(* IEC 61131-3 sources: SRCI_CLIENT_PLC/RobotLibrary/Library/POUs/Calculation/MC_CalculateTool/Structures, 4 files *)

(* ---- CalculateToolOutCmd.st ---- *)
{attribute 'pack_mode' := '1'}
// -------------------------------------------------------------------------
//  SRCI Robot Library
// -------------------------------------------------------------------------
//
//  Object:      CalculateToolOutCmd
//  Author:      Thorsten Brach
//  Date:        2024-06-09
//
//  Description:
//
//
//  Copyright:
//    (C) 2024 Thorsten Brach. All rights reserved
//             Licensed under the MIT License.
//
//  Disclaimer:
//    This project is provided without any guarantee and can be used for
//    private and commercial purposes. Any use is at the user’s
//    own risk and responsibility.
//
// -------------------------------------------------------------------------
TYPE CalculateToolOutCmd :
STRUCT
  /// Tool data
  ToolData           : ToolData;
  /// Maximum error of deviation of the TCP position
  /// from the fix point in world coordinate system
  /// If not supported: • -1
  TCPMaxError       : REAL;
  /// Average error of TCP position from the fix point  in world coordinate system
  /// If not supported: • -1
  TCPMeanError      : REAL;
END_STRUCT
END_TYPE

(* ---- CalculateToolParCmd.st ---- *)
{attribute 'pack_mode' := '1'}
// -------------------------------------------------------------------------
//  SRCI Robot Library
// -------------------------------------------------------------------------
//
//  Object:      CalculateToolParCmd
//  Author:      Thorsten Brach
//  Date:        2024-06-09
//
//  Description:
//
//
//  Copyright:
//    (C) 2024 Thorsten Brach. All rights reserved
//             Licensed under the MIT License.
//
//  Disclaimer:
//    This project is provided without any guarantee and can be used for
//    private and commercial purposes. Any use is at the user’s
//    own risk and responsibility.
//
// -------------------------------------------------------------------------
TYPE CalculateToolParCmd :
STRUCT
  /// Define which method should be used to calculate the tool frame
  Mode               : ToolCalculationMode;
  /// Index of target tool
  /// • 0: Flange (default)
  /// • 1..254: Tool frames
  ToolNo             : USINT;
  /// Index of target frame
  /// • 0: WCS (default)
  /// • 1..254: User frames
  FrameNo            : USINT;
  /// • True: Tool fixed
  /// • False: Tool on flange (default)
  ExternalTCP        : BOOL;
  /// Positions in cartesian coordinates for the tool frame calculation.
  PositionsArray     : ARRAY[0..5] OF RobotCartesianPosition;
END_STRUCT
END_TYPE

(* ---- CalculateToolRecvData.st ---- *)
{attribute 'pack_mode' := '1'}
// -------------------------------------------------------------------------
//  SRCI Robot Library
// -------------------------------------------------------------------------
//
//  Object:      CalculateToolRecvData
//  Author:      Thorsten Brach
//  Date:        2024-06-09
//
//  Description:
//
//
//  Copyright:
//    (C) 2024 Thorsten Brach. All rights reserved
//             Licensed under the MIT License.
//
//  Disclaimer:
//    This project is provided without any guarantee and can be used for
//    private and commercial purposes. Any use is at the user’s
//    own risk and responsibility.
//
// -------------------------------------------------------------------------
TYPE CalculateToolRecvData EXTENDS RspHeader :
STRUCT
  /// Maximum error of deviation of the TCP position
  /// from the fix point in world coordinate system
  /// If not supported: • -1
  TCPMaxError       : REAL;
  /// Average error of TCP position from the fix point  in world coordinate system
  /// If not supported: • -1
  TCPMeanError      : REAL;
  /// Tool data
  ToolData           : ToolData;
END_STRUCT
END_TYPE

(* ---- CalculateToolSendData.st ---- *)
{attribute 'pack_mode' := '1'}
// -------------------------------------------------------------------------
//  SRCI Robot Library
// -------------------------------------------------------------------------
//
//  Object:      CalculateToolSendData
//  Author:      Thorsten Brach
//  Date:        2024-06-09
//
//  Description:
//
//
//  Copyright:
//    (C) 2024 Thorsten Brach. All rights reserved
//             Licensed under the MIT License.
//
//  Disclaimer:
//    This project is provided without any guarantee and can be used for
//    private and commercial purposes. Any use is at the user’s
//    own risk and responsibility.
//
// -------------------------------------------------------------------------
TYPE CalculateToolSendData EXTENDS CmdHeader:
STRUCT
  DataIndex    : USINT;
  ///
  DataComplete : BYTE;
  /// Index of target tool
  /// • 0: Flange (default)
  /// • 1..254: Tool frames
  ToolNo       : USINT;
  /// Index of target frame
  /// • 0: WCS (default)
  /// • 1..254: User frames
  FrameNo      : USINT;
  /// Define which method should be used to calculate the tool frame
  Mode         : ToolCalculationMode;
  /// • True: Tool fixed
  /// • False: Tool on flange (default)
  ExternalTCP  : USINT;
  /// Positions in cartesian coordinates for the tool frame calculation.
  Position     : RobotCartesianPosition;
END_STRUCT
END_TYPE
